(* Logix 5000 project; controller TFF vendor 1 type 14 code 107 rev 33.11; software revision 33.04; part 29 of 38 *)
(* tags used below, declared in another part *)
   Address : DINT;   // Temp Address
   BufferSteps0_Prev : STRING25;
   Config : Configuration;   // Index Array used in configuration routines
   Index : DINT;   // Index
   Index2 : DINT;   // Index
   RecipeStepLog_DateTime_Empty : STRING25;   // Empty String
   RecipeStepLog_DateTime_Log : STRING25;   // Last Date Time Received from HMI
   RecipeStepLog_DateTime_Prev : STRING25;
   RecipeStepLog_Timer : TIMER;   // RecipeStepLog WatchDog Timer
   TIME : DINT[2];
   AI01 : ALIAS FOR AnalogPoint[28];
   AI02 : ALIAS FOR AnalogPoint[29];
   AI03 : ALIAS FOR AnalogPoint[30];
   AI04 : ALIAS FOR AnalogPoint[31];
   AI104 : ALIAS FOR AnalogPoint[17];
   AI201A : ALIAS FOR AnalogPoint[10];
   AI201A_SIG : ALIAS FOR DigitalPoint[90];
   AI201B : ALIAS FOR AnalogPoint[0];
   AI202 : ALIAS FOR AnalogPoint[9];
   AI203 : ALIAS FOR AnalogPoint[11];
   AI203_SIG : ALIAS FOR DigitalPoint[91];
   AI204 : ALIAS FOR AnalogPoint[12];
   AI204_SIG : ALIAS FOR DigitalPoint[92];
   AlarmAnalog : AlarmAnalog[50];   // Analog Alarm Array
   AlarmControl : AlarmControl;   // Alarm Control
   AlarmDeviation : AlarmDeviation[20];   // Control Loop Deviation Alarm Array
   AnalogOutput : AnalogOutput[25];   // Analog Output Array
   AnalogPoint : AnalogInput[50];   // Analog Input Array
   CCPSystem : CCPSystem;   // CCP System Data
   CPU_Scanning : BOOL;   // System Scanning Flag
   DigitalOutput : BOOL[256];   // Digital Output Array these bits are sent to output cards.
   DigitalPoint : DigitalPoint[150];   // Digital Point Array
   FI101 : ALIAS FOR AnalogPoint[19];
   FI201 : ALIAS FOR AnalogPoint[2];
   FI201_SIG : ALIAS FOR DigitalPoint[93];
   FI401 : ALIAS FOR AnalogPoint[20];
   FI401_SIG : ALIAS FOR DigitalPoint[94];
   Gateway : Gateway;   // Gateway Control
   GWModbus : IO_Station;   // Status of Gateway Modbus
   HTCCollectorError : BOOL;   // Historical Data Collector Error (Set to 1 by HMI if Error)
   HTCHeartBeat : BOOL;   // Historical Data Collection heartbeat (Set to 1 by HMI Reset to 0 by PLC)
   MIX101 : ALIAS FOR AnalogPoint[14];
   Mixer : Mixer;   // Mixer config. structure
   OperatingTime : OperatingTime;
   PcToPLCHeartBeat : BOOL;   // PC to PLC communication heartbeat Set to 1 by HMI Reset to 0 by plc
   PCV101 : ALIAS FOR AnalogPoint[3];
   PCV201 : ALIAS FOR AnalogPoint[4];
   Phase0 : ALIAS FOR Phase[0];   // Phase 0
   PI001 : ALIAS FOR AnalogPoint[5];
   PI001_SIG : ALIAS FOR DigitalPoint[97];
   PI101 : ALIAS FOR AnalogPoint[6];
   PI201 : ALIAS FOR AnalogPoint[7];
   PI401 : ALIAS FOR AnalogPoint[8];
   PI601 : ALIAS FOR AnalogPoint[21];
   PI601_SIG : ALIAS FOR DigitalPoint[95];
   PLCFault : FaultRecordType;   // PLC Major Fault Record
   Rack_ACT350_WI101_200L : IO_Station;   // Status of ACT350 200L
   Rack_ACT350_WI101_500L : IO_Station;   // Status of ACT350 500L
   Rack_Murr_Node0_Smart : IO_Station;   // Status of Node 0 Smart
   Rack_Murr_Node1_TFF20 : IO_Station;   // Status of Node 1 TFF20
   Rack_Murr_Node1_TFF40 : IO_Station;   // Status of Node 1 TFF40
   Rack_Murr_Node1_TFF80 : IO_Station;   // Status of Node 1 TFF80
   RawAnalogInputArray : INT[50];   // Array of analog input raw
   RecipeStepLog_DateTime : STRING25;
   SysControl : SysControl;   // General system status and command
   Tank : TankManagement;   // Tank Management
   TCU101 : ALIAS FOR AnalogPoint[18];
   ThisSystem : SystemType;
   TI101 : ALIAS FOR AnalogPoint[13];
   TI201 : ALIAS FOR AnalogPoint[22];
   WI201 : ALIAS FOR AnalogPoint[1];
   WI201_SIG : ALIAS FOR DigitalPoint[96];
   XS011 : ALIAS FOR DigitalPoint[14];
   XS012 : ALIAS FOR DigitalPoint[15];
   YA01 : ALIAS FOR DigitalPoint[50];
   YA02 : ALIAS FOR DigitalPoint[51];
   YA03 : ALIAS FOR DigitalPoint[52];
   YA06 : ALIAS FOR DigitalPoint[55];
   YA07 : ALIAS FOR DigitalPoint[56];
   YA08 : ALIAS FOR DigitalPoint[57];
   YA09 : ALIAS FOR DigitalPoint[58];
   YA10 : ALIAS FOR DigitalPoint[59];
   YA13 : ALIAS FOR DigitalPoint[62];
   YA14 : ALIAS FOR DigitalPoint[63];
   YA15 : ALIAS FOR DigitalPoint[69];
   YA16 : ALIAS FOR DigitalPoint[70];
   YA17 : ALIAS FOR DigitalPoint[71];
   YA18 : ALIAS FOR DigitalPoint[72];
   YA41 : ALIAS FOR DigitalPoint[73];
   ZS001 : ALIAS FOR DigitalPoint[6];
   ZS002 : ALIAS FOR DigitalPoint[7];
   ZS003 : ALIAS FOR DigitalPoint[8];
   ZS004 : ALIAS FOR DigitalPoint[9];
   ZS005 : ALIAS FOR DigitalPoint[10];
   ZSDF : ALIAS FOR DigitalPoint[68];
(* Process, continued *)

ROUTINE FaultRoutine   (* ladder *)
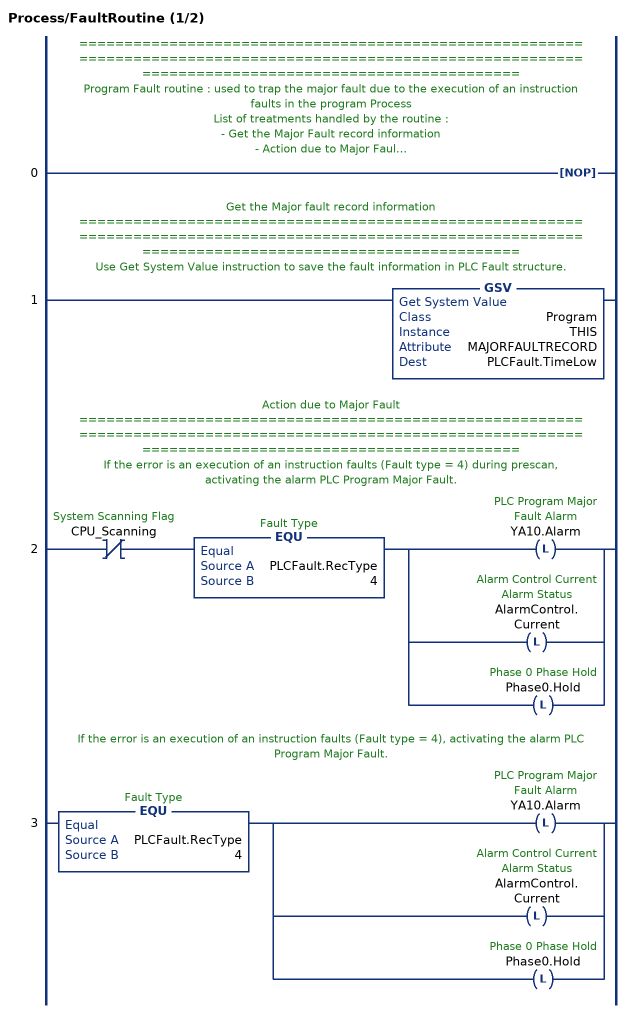
   // ==========================================================================================================================================================
   //                                                               Program Fault routine : used to trap the major fault due to the execution of an instruction faults in the program Process
   //                                                     List of treatments handled by the routine :
   //                                                          - Get the Major Fault record information
   //                                                          - Action due to Major Fault
   //                                                     -----------------------------------------------------------------------------------------------------------------------------------------------------
   //                                                     History
   // 		2019-DEC-24 - Merck - Q. Spindler - Initial version for Candidate Release 1.00.00.00.a
   // ==========================================================================================================================================================
   0: NOP();
   // Get the Major fault record information
   // ==========================================================================================================================================================
   // Use Get System Value instruction to save the fault information in PLC Fault structure.
   1: GSV(Program,THIS,MAJORFAULTRECORD,PLCFault.TimeLow);
   // Action due to Major Fault
   // ==========================================================================================================================================================
   // If the error is an execution of an instruction faults (Fault type = 4) during prescan, activating the alarm PLC Program Major Fault.
   2: XIO(CPU_Scanning)EQU(PLCFault.RecType,4)[OTL(YA10.Alarm) ,OTL(AlarmControl.Current) ,OTL(Phase0.Hold) ];
   // If the error is an execution of an instruction faults (Fault type = 4), activating the alarm PLC Program Major Fault.
   3: EQU(PLCFault.RecType,4)[OTL(YA10.Alarm) ,OTL(AlarmControl.Current) ,OTL(Phase0.Hold) ];
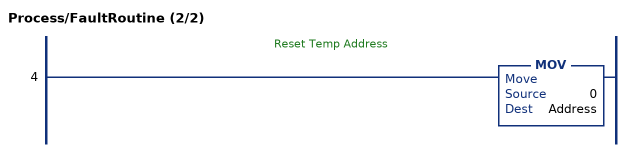
   // Reset Temp Address
   4: MOV(0,Address);
END_ROUTINE

ROUTINE Gateway   (* structured text *)
   (* ==========================================================
   	Gateway : Mapping Data to gateway communication Table
   		format of data transfered is DINT.
   		REAL type Data (Analog) must managed to convert it to DINT format with an accuracy of 3 digits (x1000 for Data sended, /1000 for Data received.
   
   	List of treatments
   		- Write to the gateway
   		- Read from the gateway
   		- Gateway wattchdog  processing
   
   -----------------------------------------------------------------------------------------------------------------------------------------------------
   	History
   		2019-DEC-24 - Merck - Q. Spindler - Initial version for Candidate Release 1.00.00.00.a
   		2020-MAR-25 - Merck - Q. Spindler - Modifications for Candidate Release 1.00.00.00.b
   					- Change Analog output indexes that caused PLC major Fault
   ============================================================*)
   
   
   
   (* Write to the gateway
   =========================================================================*)
   
   (* Send analog Point to the gateway*)
   FOR Gateway.Index := 0 TO 46 BY 1 DO
   	Gateway.Output[Gateway.Index]:= AnalogPoint[Gateway.Index].CurrentValue*1000;
   END_FOR;
   
   (* Send analog output to the gateway*)
   FOR Gateway.Index := 47 TO 58 BY 1 DO
   	Gateway.Output[Gateway.Index]:= AnalogOutput[Gateway.Index-47].ScaledValue*1000;
   END_FOR;
   
   (* Send Digital Point to the gateway*)
   FOR Gateway.Index := 0 TO 31 BY 1 DO
   	Gateway.Output[59].[Gateway.Index]:= DigitalPoint[Gateway.Index].CurrentValue;
   	Gateway.Output[60].[Gateway.Index]:= DigitalPoint[Gateway.Index+32].CurrentValue;
   	Gateway.Output[61].[Gateway.Index]:= DigitalPoint[Gateway.Index+50].SoftInput;
   	Gateway.Output[62].[Gateway.Index]:= DigitalPoint[Gateway.Index+82].SoftInput;
   END_FOR;
   
   (* Send Digital Output to the gateway *)
   FOR Gateway.Index := 0 TO 31 BY 1 DO
   	Gateway.Output[63].[Gateway.Index]:= DigitalOutput[Gateway.Index];
   	Gateway.Output[64].[Gateway.Index]:= DigitalOutput[Gateway.Index+32];
   	Gateway.Output[65].[Gateway.Index]:= DigitalOutput[Gateway.Index+64];
   END_FOR;
   
   (* Send Digital Alarm to the gateway*)
   FOR Gateway.Index := 0 TO 31 BY 1 DO
   	Gateway.Output[66].[Gateway.Index]:= DigitalPoint[Gateway.Index].Alarm;
   	Gateway.Output[67].[Gateway.Index]:= DigitalPoint[Gateway.Index+32].Alarm;
   	Gateway.Output[68].[Gateway.Index]:= DigitalPoint[Gateway.Index+64].Alarm;
   	Gateway.Output[69].[Gateway.Index]:= DigitalPoint[Gateway.Index+96].Alarm;
   END_FOR;
   
   
   (* Send Analog Alarm to the gateway*)
   FOR Gateway.Index := 70 TO 75 BY 1 DO
   	FOR Gateway.Index2 := 0 TO 31 BY 4 DO
   		Gateway.Output[Gateway.Index].[Gateway.Index2] := AlarmAnalog[(Gateway.Index2 / 4)+((Gateway.Index-70) * 8)].LOLOAlarm;
   		Gateway.Output[Gateway.Index].[Gateway.Index2 + 1] := AlarmAnalog[(Gateway.Index2 / 4)+((Gateway.Index-70) * 8)].LOAlarm;
   		Gateway.Output[Gateway.Index].[Gateway.Index2 + 2] := AlarmAnalog[(Gateway.Index2 / 4)+((Gateway.Index-70) * 8)].HIAlarm;
   		Gateway.Output[Gateway.Index].[Gateway.Index2 + 3] := AlarmAnalog[(Gateway.Index2 / 4)+((Gateway.Index-70) * 8)].HIHIAlarm;
   	END_FOR;
   END_FOR;
   
   
   (* Send Deviqtions Alarm to the gateway*)
   FOR Gateway.Index := 0 TO 15 BY 1 DO
   	Gateway.Output[76].[Gateway.Index * 2] := AlarmDeviation[Gateway.Index].HIAlarm;
   	Gateway.Output[76].[Gateway.Index * 2 + 1] := AlarmDeviation[Gateway.Index].HIHIAlarm;
   END_FOR;
   
   (* Clear unused space*)
   FOR Gateway.Index := 77 TO 81 BY 1 DO
   	Gateway.Output[Gateway.Index] := 0;
   END_FOR;
   
   
   (* Send CCP System status, system in alarm status, system in maintenance mode status to the gateway*)
   Gateway.Output[82] := CCPSystem.State;
   Gateway.Output[83].0 := AlarmControl.AlarmHigh ;
   Gateway.Output[83].1 := AlarmControl.AlarmLow ;
   Gateway.Output[83].2 := SysControl.Maintenance;
   
   (* Send Analog Action from recipe to the gateway *)
   FOR Gateway.Index := 84 TO 103 BY 1 DO
   	Gateway.Output[Gateway.Index]:= Gateway.RecipeAction_Analog[Gateway.Index-84]*1000;
   END_FOR;
   
   (* Send Digital Action from recipe to the gateway *)
   FOR Gateway.Index := 104 TO 105 BY 1 DO
   	Gateway.Output[Gateway.Index]:= Gateway.RecipeAction_Digital[Gateway.Index-104];
   END_FOR;
   
   (* Send Watchdog data to the gateway *)
   Gateway.Output[106] := Gateway.Watchdog_Out_Skid;
   Gateway.Output[107] := Gateway.Watchdog_Out_Ext;
   
   (* Data Send to the Gateway*)
   FOR Gateway.Index := 0 TO 123 BY 1 DO
   	GATEWAY:O.Data[Gateway.Index] := Gateway.Output[Gateway.Index];
   END_FOR;
   
   
   (* Read from the gateway
   =========================================================================*)
   
   (* Read from the gateway tha analog criteria for recipe *)
   FOR Gateway.Index := 0 TO 19 BY 1 DO
   		Gateway.RecipeCriteria_Analog[Gateway.Index] := Gateway.Input[Gateway.Index]/1000;
   END_FOR;
   
   (* Read from the gateway tha digital criteria for recipe *)
   FOR Gateway.Index := 20 TO 21 BY 1 DO
   		Gateway.RecipeCriteria_Digital[Gateway.Index-20] := Gateway.Input[Gateway.Index];
   END_FOR;
   
   (* Read Watchdog data from the gateway *)
   Gateway.Watchdog_In_Skid := Gateway.Input[22];
   Gateway.Watchdog_In_Ext := Gateway.Input[23];
   
   (* Data receive from the Gateway *)
   FOR Gateway.Index := 0 TO 63 BY 1 DO
   	Gateway.Input[Gateway.Index] := GATEWAY:I.Data[Gateway.Index];
   END_FOR;
   
   
   
   (* Gateway wattchdog  processing
   =========================================================================*)
   
   (* Verify if skid watchdog value receive is equal to watchdog value send previously *)
   IF Gateway.Watchdog_Out_Skid = Gateway.Watchdog_In_Skid Then
   	(* Add 1 to skid watchdog value *)
   	Gateway.Watchdog_Out_Skid := Gateway.Watchdog_Out_Skid +1;
   	(* Set to 1 YA16 soft input (alarm watchdog) *)
   	YA16.SoftInput := 1 ;
   Else
   	(* Set to 0 YA16 soft input (alarm watchdog) *)
   	YA16.SoftInput := 0 ;
   End_If;
   
   (* If skid watchdog value is greater than 9999, reset value *)
   IF Gateway.Watchdog_Out_Skid > 9999 Then
   	Gateway.Watchdog_Out_Skid := 0;
   End_IF;
   
   (* Copy external watchdog value received in the one to be sent *)
   Gateway.Watchdog_Out_Ext := Gateway.Watchdog_In_Ext;
END_ROUTINE

ROUTINE InputAnalogPoint   (* ladder *)
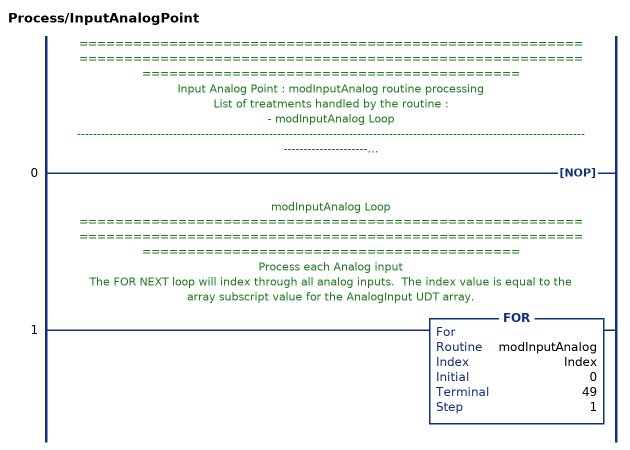
   // ==========================================================================================================================================================
   //                                                                                                             Input Analog Point : modInputAnalog routine processing
   //                                                     List of treatments handled by the routine :
   //                                                          - modInputAnalog Loop
   //                                                     -----------------------------------------------------------------------------------------------------------------------------------------------------
   //                                                     History
   // 		2019-DEC-24 - Merck - Q. Spindler - Initial version for Candidate Release 1.00.00.00.a
   // ==========================================================================================================================================================
   0: NOP();
   // modInputAnalog Loop
   // ==========================================================================================================================================================
   // Process each Analog input
   // The FOR NEXT loop will index through all analog inputs.  The index value is equal to the array subscript value for the AnalogInput UDT array.
   1: FOR(modInputAnalog,Index,0,49,1);
END_ROUTINE

ROUTINE InputAnalogRaw   (* ladder *)
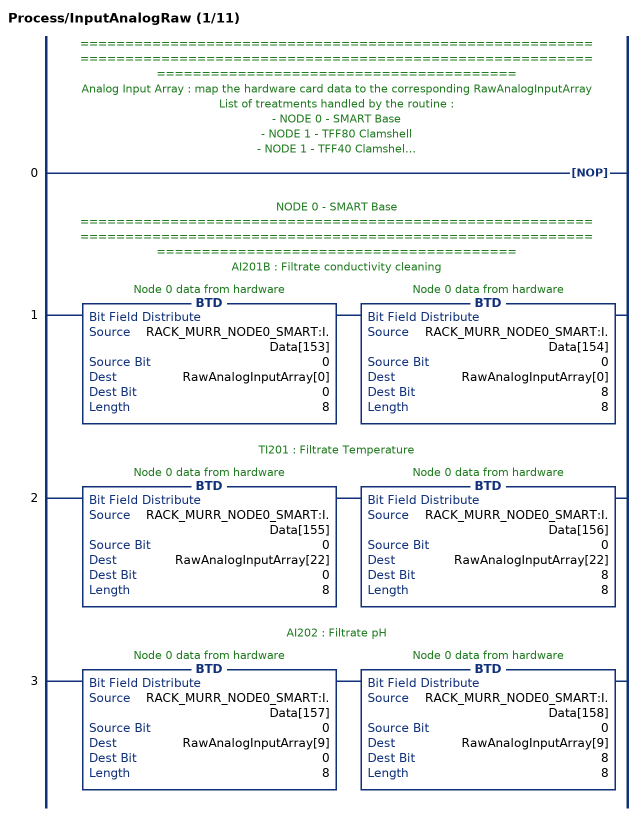
   // ==========================================================================================================================================================
   //                                                                                          Analog Input Array : map the hardware card data to the corresponding RawAnalogInputArray
   //                                                     List of treatments handled by the routine :
   //                                                    - NODE 0 - SMART Base
   //                                                         - NODE 1 - TFF80 Clamshell
   //                                                         - NODE 1 - TFF40 Clamshell
   //                                                         - NODE 1 - TFF20 Clamshell
   //                                                     -----------------------------------------------------------------------------------------------------------------------------------------------------
   //                                                     History
   // 		2019-DEC-24 - Merck - Q. Spindler - Initial version for Candidate Release 1.00.00.00.a
   //                                 2020-APR-09 - Merck - Q. Spindler - Modifications for Candidate Release 1.00.00.00.b
   //                  - Change IO address for MIX101
   //                                 2022-SEP-28 - Actemium - J. Jaekel - Modifications for Candidate Release 1.01.00.01.a
   // - Add TI201
   // ==========================================================================================================================================================
   0: NOP();
   // NODE 0 - SMART Base
   // ==========================================================================================================================================================
   // AI201B : Filtrate conductivity cleaning
   1: BTD(RACK_MURR_NODE0_SMART:I.Data[153],0,RawAnalogInputArray[0],0,8)BTD(RACK_MURR_NODE0_SMART:I.Data[154],0,RawAnalogInputArray[0],8,8);
   // TI201 : Filtrate Temperature
   2: BTD(RACK_MURR_NODE0_SMART:I.Data[155],0,RawAnalogInputArray[22],0,8)BTD(RACK_MURR_NODE0_SMART:I.Data[156],0,RawAnalogInputArray[22],8,8);
   // AI202 : Filtrate pH
   3: BTD(RACK_MURR_NODE0_SMART:I.Data[157],0,RawAnalogInputArray[9],0,8)BTD(RACK_MURR_NODE0_SMART:I.Data[158],0,RawAnalogInputArray[9],8,8);
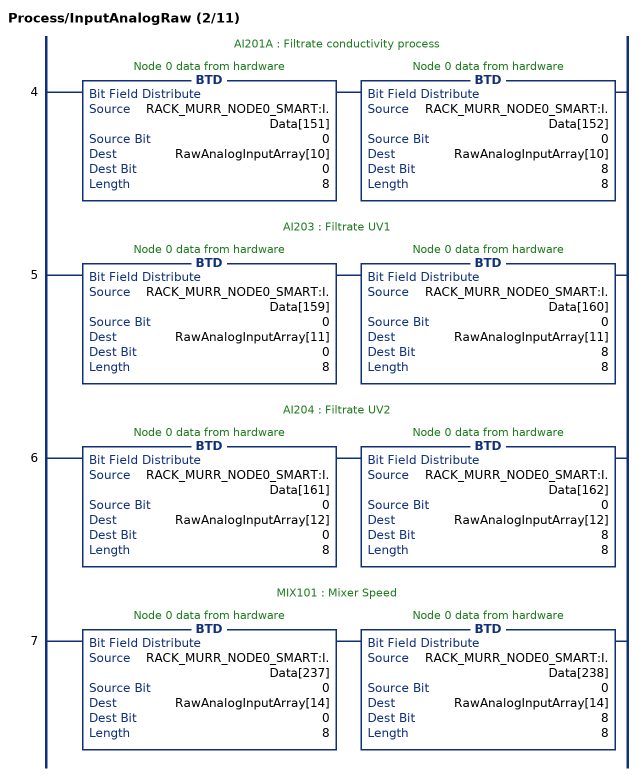
   // AI201A : Filtrate conductivity process
   4: BTD(RACK_MURR_NODE0_SMART:I.Data[151],0,RawAnalogInputArray[10],0,8)BTD(RACK_MURR_NODE0_SMART:I.Data[152],0,RawAnalogInputArray[10],8,8);
   // AI203 : Filtrate UV1
   5: BTD(RACK_MURR_NODE0_SMART:I.Data[159],0,RawAnalogInputArray[11],0,8)BTD(RACK_MURR_NODE0_SMART:I.Data[160],0,RawAnalogInputArray[11],8,8);
   // AI204 : Filtrate UV2
   6: BTD(RACK_MURR_NODE0_SMART:I.Data[161],0,RawAnalogInputArray[12],0,8)BTD(RACK_MURR_NODE0_SMART:I.Data[162],0,RawAnalogInputArray[12],8,8);
   // MIX101 : Mixer Speed
   7: BTD(RACK_MURR_NODE0_SMART:I.Data[237],0,RawAnalogInputArray[14],0,8)BTD(RACK_MURR_NODE0_SMART:I.Data[238],0,RawAnalogInputArray[14],8,8);
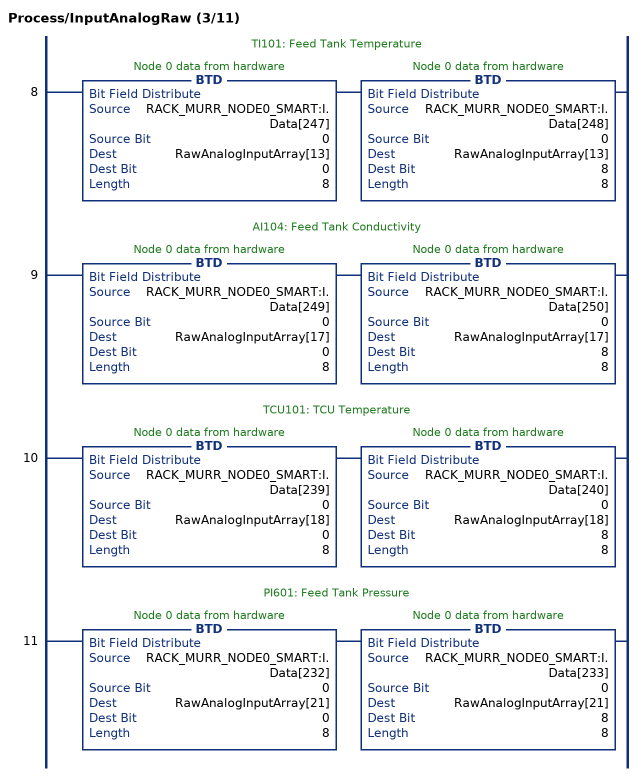
   // TI101: Feed Tank Temperature
   8: BTD(RACK_MURR_NODE0_SMART:I.Data[247],0,RawAnalogInputArray[13],0,8)BTD(RACK_MURR_NODE0_SMART:I.Data[248],0,RawAnalogInputArray[13],8,8);
   // AI104: Feed Tank Conductivity
   9: BTD(RACK_MURR_NODE0_SMART:I.Data[249],0,RawAnalogInputArray[17],0,8)BTD(RACK_MURR_NODE0_SMART:I.Data[250],0,RawAnalogInputArray[17],8,8);
   // TCU101: TCU Temperature
   10: BTD(RACK_MURR_NODE0_SMART:I.Data[239],0,RawAnalogInputArray[18],0,8)BTD(RACK_MURR_NODE0_SMART:I.Data[240],0,RawAnalogInputArray[18],8,8);
   // PI601: Feed Tank Pressure
   11: BTD(RACK_MURR_NODE0_SMART:I.Data[232],0,RawAnalogInputArray[21],0,8)BTD(RACK_MURR_NODE0_SMART:I.Data[233],0,RawAnalogInputArray[21],8,8);
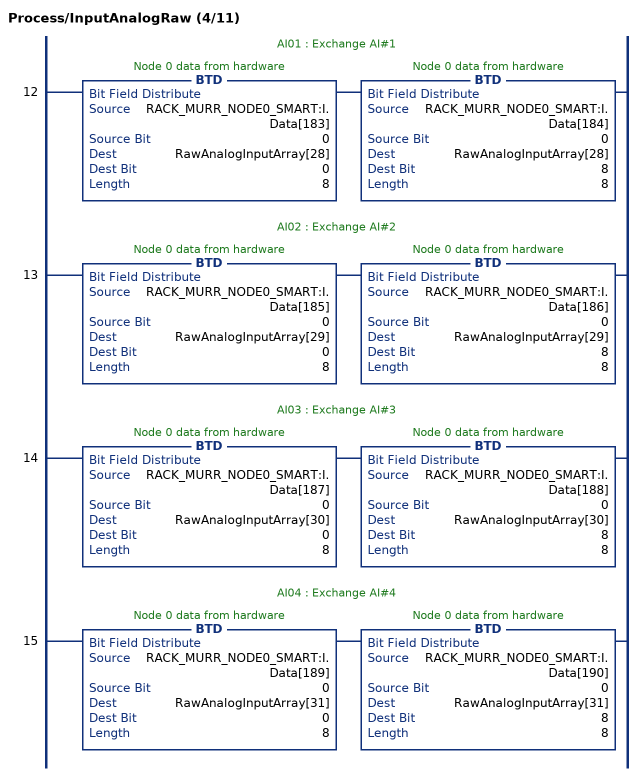
   // AI01 : Exchange AI#1
   12: BTD(RACK_MURR_NODE0_SMART:I.Data[183],0,RawAnalogInputArray[28],0,8)BTD(RACK_MURR_NODE0_SMART:I.Data[184],0,RawAnalogInputArray[28],8,8);
   // AI02 : Exchange AI#2
   13: BTD(RACK_MURR_NODE0_SMART:I.Data[185],0,RawAnalogInputArray[29],0,8)BTD(RACK_MURR_NODE0_SMART:I.Data[186],0,RawAnalogInputArray[29],8,8);
   // AI03 : Exchange AI#3
   14: BTD(RACK_MURR_NODE0_SMART:I.Data[187],0,RawAnalogInputArray[30],0,8)BTD(RACK_MURR_NODE0_SMART:I.Data[188],0,RawAnalogInputArray[30],8,8);
   // AI04 : Exchange AI#4
   15: BTD(RACK_MURR_NODE0_SMART:I.Data[189],0,RawAnalogInputArray[31],0,8)BTD(RACK_MURR_NODE0_SMART:I.Data[190],0,RawAnalogInputArray[31],8,8);
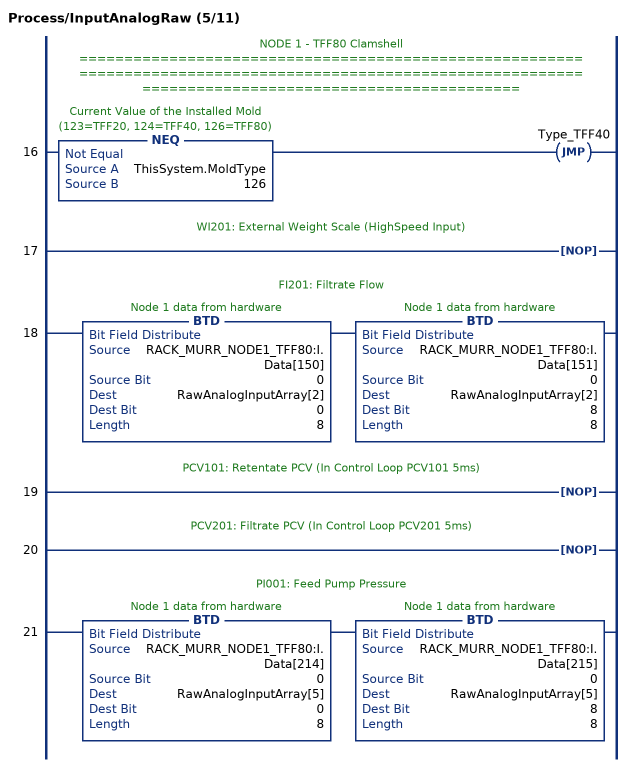
   // NODE 1 - TFF80 Clamshell
   // ==========================================================================================================================================================
   16: NEQ(ThisSystem.MoldType,126)JMP(Type_TFF40);
   // WI201: External Weight Scale (HighSpeed Input)
   17: NOP();
   // FI201: Filtrate Flow
   18: BTD(RACK_MURR_NODE1_TFF80:I.Data[150],0,RawAnalogInputArray[2],0,8)BTD(RACK_MURR_NODE1_TFF80:I.Data[151],0,RawAnalogInputArray[2],8,8);
   // PCV101: Retentate PCV (In Control Loop PCV101 5ms)
   19: NOP();
   // PCV201: Filtrate PCV (In Control Loop PCV201 5ms)
   20: NOP();
   // PI001: Feed Pump Pressure
   21: BTD(RACK_MURR_NODE1_TFF80:I.Data[214],0,RawAnalogInputArray[5],0,8)BTD(RACK_MURR_NODE1_TFF80:I.Data[215],0,RawAnalogInputArray[5],8,8);
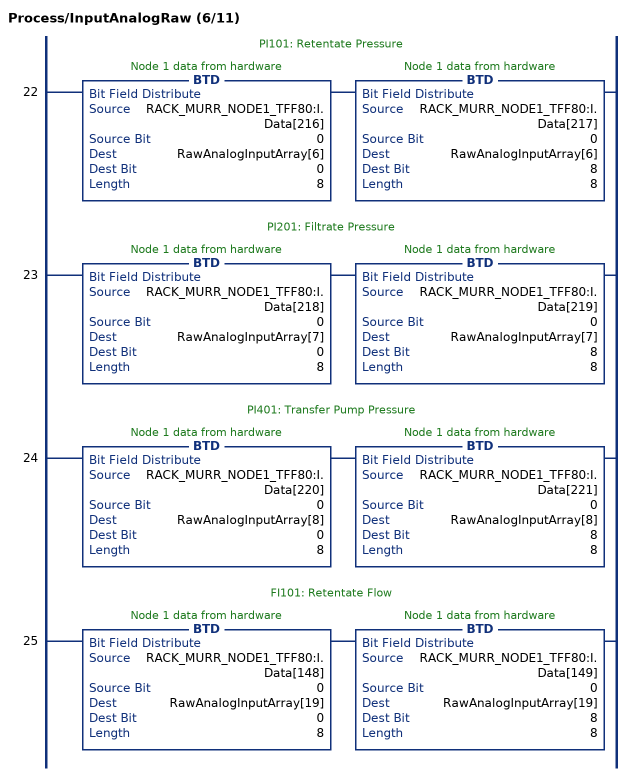
   // PI101: Retentate Pressure
   22: BTD(RACK_MURR_NODE1_TFF80:I.Data[216],0,RawAnalogInputArray[6],0,8)BTD(RACK_MURR_NODE1_TFF80:I.Data[217],0,RawAnalogInputArray[6],8,8);
   // PI201: Filtrate Pressure
   23: BTD(RACK_MURR_NODE1_TFF80:I.Data[218],0,RawAnalogInputArray[7],0,8)BTD(RACK_MURR_NODE1_TFF80:I.Data[219],0,RawAnalogInputArray[7],8,8);
   // PI401: Transfer Pump Pressure
   24: BTD(RACK_MURR_NODE1_TFF80:I.Data[220],0,RawAnalogInputArray[8],0,8)BTD(RACK_MURR_NODE1_TFF80:I.Data[221],0,RawAnalogInputArray[8],8,8);
   // FI101: Retentate Flow
   25: BTD(RACK_MURR_NODE1_TFF80:I.Data[148],0,RawAnalogInputArray[19],0,8)BTD(RACK_MURR_NODE1_TFF80:I.Data[149],0,RawAnalogInputArray[19],8,8);
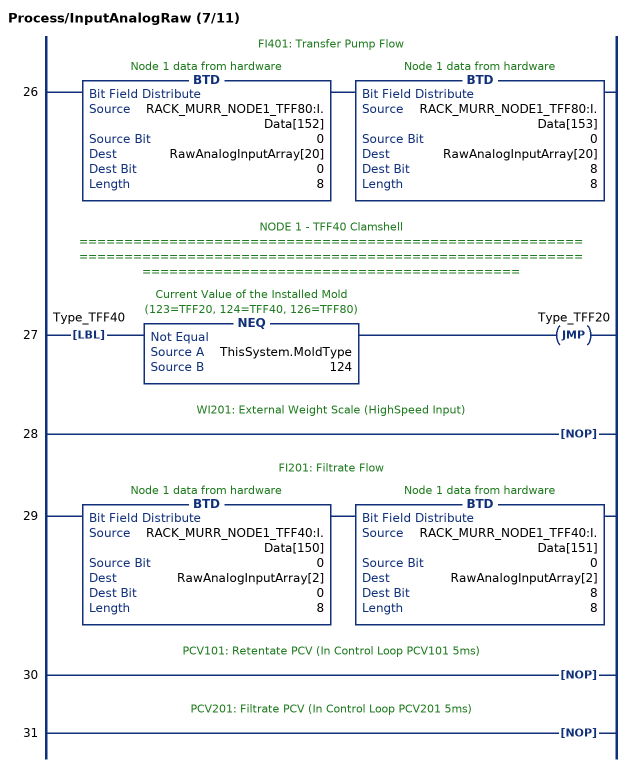
   // FI401: Transfer Pump Flow
   26: BTD(RACK_MURR_NODE1_TFF80:I.Data[152],0,RawAnalogInputArray[20],0,8)BTD(RACK_MURR_NODE1_TFF80:I.Data[153],0,RawAnalogInputArray[20],8,8);
   // NODE 1 - TFF40 Clamshell
   // ==========================================================================================================================================================
   27: LBL(Type_TFF40)NEQ(ThisSystem.MoldType,124)JMP(Type_TFF20);
   // WI201: External Weight Scale (HighSpeed Input)
   28: NOP();
   // FI201: Filtrate Flow
   29: BTD(RACK_MURR_NODE1_TFF40:I.Data[150],0,RawAnalogInputArray[2],0,8)BTD(RACK_MURR_NODE1_TFF40:I.Data[151],0,RawAnalogInputArray[2],8,8);
   // PCV101: Retentate PCV (In Control Loop PCV101 5ms)
   30: NOP();
   // PCV201: Filtrate PCV (In Control Loop PCV201 5ms)
   31: NOP();
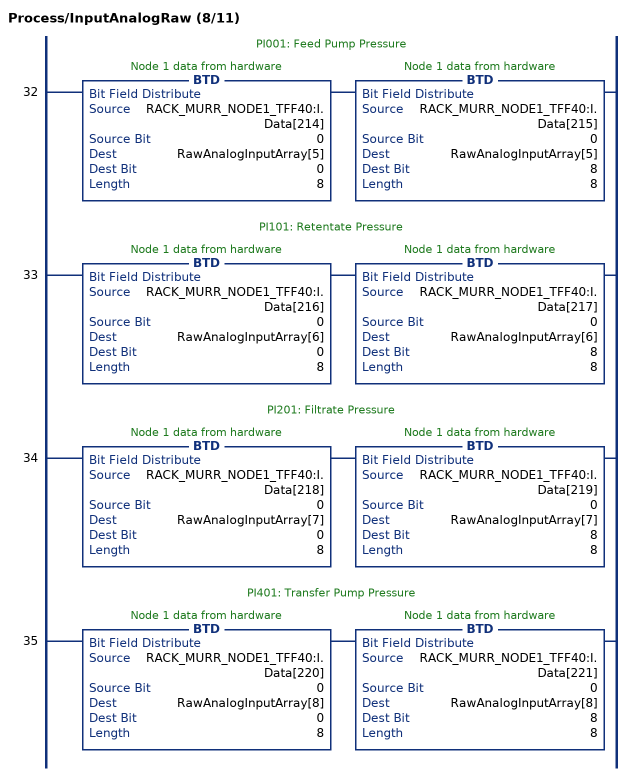
   // PI001: Feed Pump Pressure
   32: BTD(RACK_MURR_NODE1_TFF40:I.Data[214],0,RawAnalogInputArray[5],0,8)BTD(RACK_MURR_NODE1_TFF40:I.Data[215],0,RawAnalogInputArray[5],8,8);
   // PI101: Retentate Pressure
   33: BTD(RACK_MURR_NODE1_TFF40:I.Data[216],0,RawAnalogInputArray[6],0,8)BTD(RACK_MURR_NODE1_TFF40:I.Data[217],0,RawAnalogInputArray[6],8,8);
   // PI201: Filtrate Pressure
   34: BTD(RACK_MURR_NODE1_TFF40:I.Data[218],0,RawAnalogInputArray[7],0,8)BTD(RACK_MURR_NODE1_TFF40:I.Data[219],0,RawAnalogInputArray[7],8,8);
   // PI401: Transfer Pump Pressure
   35: BTD(RACK_MURR_NODE1_TFF40:I.Data[220],0,RawAnalogInputArray[8],0,8)BTD(RACK_MURR_NODE1_TFF40:I.Data[221],0,RawAnalogInputArray[8],8,8);
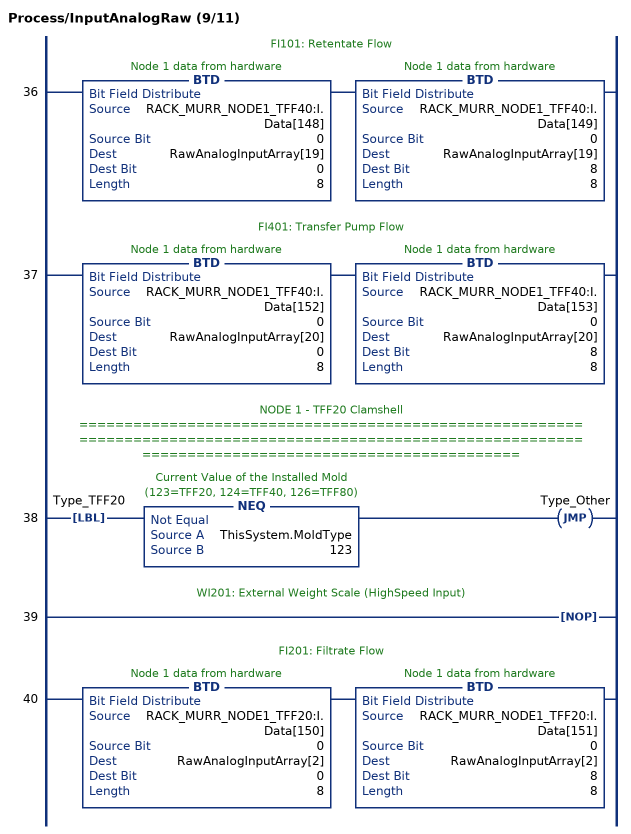
   // FI101: Retentate Flow
   36: BTD(RACK_MURR_NODE1_TFF40:I.Data[148],0,RawAnalogInputArray[19],0,8)BTD(RACK_MURR_NODE1_TFF40:I.Data[149],0,RawAnalogInputArray[19],8,8);
   // FI401: Transfer Pump Flow
   37: BTD(RACK_MURR_NODE1_TFF40:I.Data[152],0,RawAnalogInputArray[20],0,8)BTD(RACK_MURR_NODE1_TFF40:I.Data[153],0,RawAnalogInputArray[20],8,8);
   // NODE 1 - TFF20 Clamshell
   // ==========================================================================================================================================================
   38: LBL(Type_TFF20)NEQ(ThisSystem.MoldType,123)JMP(Type_Other);
   // WI201: External Weight Scale (HighSpeed Input)
   39: NOP();
   // FI201: Filtrate Flow
   40: BTD(RACK_MURR_NODE1_TFF20:I.Data[150],0,RawAnalogInputArray[2],0,8)BTD(RACK_MURR_NODE1_TFF20:I.Data[151],0,RawAnalogInputArray[2],8,8);
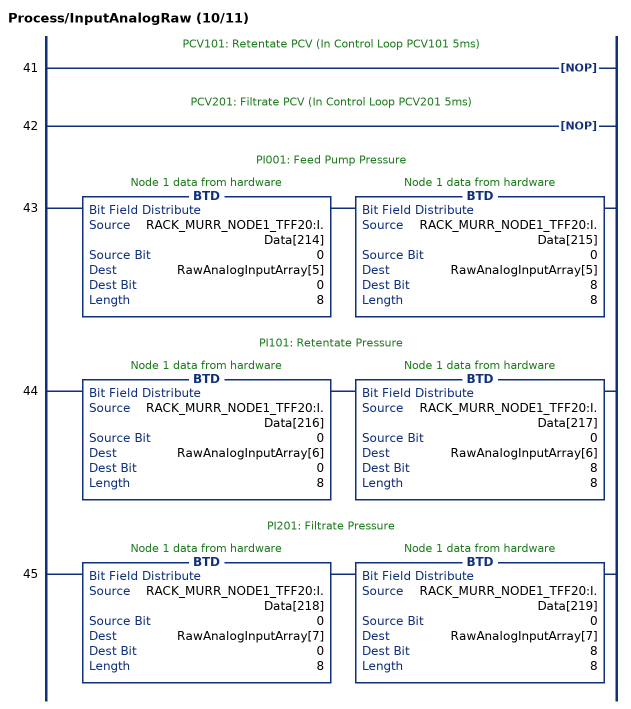
   // PCV101: Retentate PCV (In Control Loop PCV101 5ms)
   41: NOP();
   // PCV201: Filtrate PCV (In Control Loop PCV201 5ms)
   42: NOP();
   // PI001: Feed Pump Pressure
   43: BTD(RACK_MURR_NODE1_TFF20:I.Data[214],0,RawAnalogInputArray[5],0,8)BTD(RACK_MURR_NODE1_TFF20:I.Data[215],0,RawAnalogInputArray[5],8,8);
   // PI101: Retentate Pressure
   44: BTD(RACK_MURR_NODE1_TFF20:I.Data[216],0,RawAnalogInputArray[6],0,8)BTD(RACK_MURR_NODE1_TFF20:I.Data[217],0,RawAnalogInputArray[6],8,8);
   // PI201: Filtrate Pressure
   45: BTD(RACK_MURR_NODE1_TFF20:I.Data[218],0,RawAnalogInputArray[7],0,8)BTD(RACK_MURR_NODE1_TFF20:I.Data[219],0,RawAnalogInputArray[7],8,8);
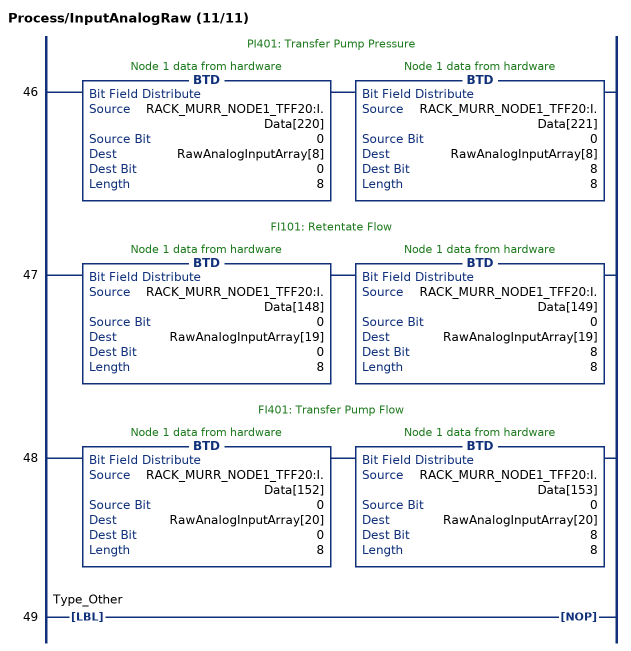
   // PI401: Transfer Pump Pressure
   46: BTD(RACK_MURR_NODE1_TFF20:I.Data[220],0,RawAnalogInputArray[8],0,8)BTD(RACK_MURR_NODE1_TFF20:I.Data[221],0,RawAnalogInputArray[8],8,8);
   // FI101: Retentate Flow
   47: BTD(RACK_MURR_NODE1_TFF20:I.Data[148],0,RawAnalogInputArray[19],0,8)BTD(RACK_MURR_NODE1_TFF20:I.Data[149],0,RawAnalogInputArray[19],8,8);
   // FI401: Transfer Pump Flow
   48: BTD(RACK_MURR_NODE1_TFF20:I.Data[152],0,RawAnalogInputArray[20],0,8)BTD(RACK_MURR_NODE1_TFF20:I.Data[153],0,RawAnalogInputArray[20],8,8);
   49: LBL(Type_Other)NOP();
END_ROUTINE

ROUTINE InputDigitalPoint   (* ladder *)
// Digital Point Routine
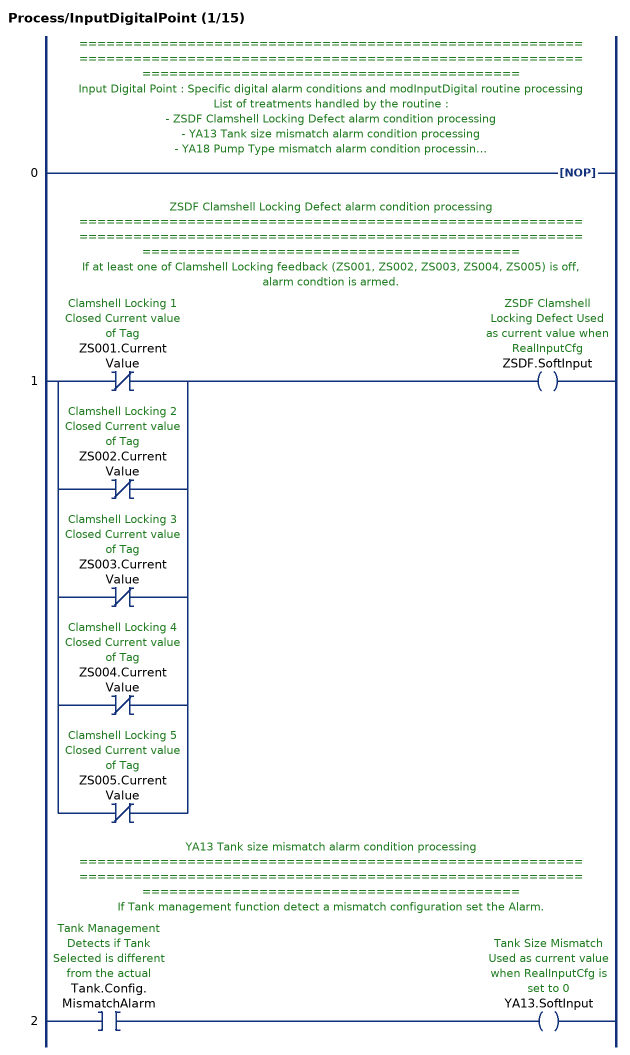
   // ==========================================================================================================================================================
   //                                                                                   Input Digital Point : Specific digital alarm conditions and modInputDigital routine processing
   //                                                     List of treatments handled by the routine :
   //                                                          - ZSDF Clamshell Locking Defect alarm condition processing
   //                                                          - YA13 Tank size mismatch alarm condition processing
   //                                                          - YA18 Pump Type mismatch alarm condition processing
   //                                                          - YA03 Historical data collection failure alarm condition processing
   //                                                          - YA01 PC to PLC com. failure alarm condition processing
   //                                                          - YA02 CCP Runtime com. failure alarm condition processing
   //                                                          - YA14 SQL Write failure alarm condition processing
   //                                                          - Node 0 communication failure and internal defect (YA06 and YA07)
   //                                                          - Node 1 communication failure and internal defect (YA08 and YA09)
   //                                                          - ACT350 communication failure (YA15)
   //                                                          - Operating Time Exceeded (YA41)
   //                                                          - Analog Signal Failure
   //                                                          - modInputDigital Loop
   //                                                     -----------------------------------------------------------------------------------------------------------------------------------------------------
   //                                                     History
   // 		2019-DEC-24 - Merck - Q. Spindler - Initial version for Candidate Release 1.00.00.00.a
   // 		2020-APR-06 - Merck - Q. Spindler - Modifications for Candidate Release 1.00.00.00.b
   //                                                             - Trigger pressure signal failure when the raw value equal to the RawMax
   // 		2020-JUN-09 - Merck - Q. Spindler - Modifications for Candidate Release 1.00.00.00.c
   //                                                             - Change Alarm condition for YA07 and YA09, internal defect dont trigger if the Node is not connected
   // - Change YA14 Alarm condition processing to add HMI Watchdog
   // 		2021-OCT-26 - Merck - Q. Spindler - Modifications for Candidate Release 1.01.00.00.a
   // - Add HTC Collector Error in the YA03 alarm conditions
   //   - Add Operating Time Exceeded (YA41)
   // 		2022-SEP-26 - Actemium - J. Jaekel - Modifications for Candidate Release 1.01.00.01.a
   // - Add TI201 signal failure
   // ==========================================================================================================================================================
   0: NOP();
   // ZSDF Clamshell Locking Defect alarm condition processing
   // ==========================================================================================================================================================
   // If at least one of Clamshell Locking feedback (ZS001, ZS002, ZS003, ZS004, ZS005) is off, alarm condtion is armed.
   1: [XIO(ZS001.CurrentValue) ,XIO(ZS002.CurrentValue) ,XIO(ZS003.CurrentValue) ,XIO(ZS004.CurrentValue) ,XIO(ZS005.CurrentValue) ]OTE(ZSDF.SoftInput);
   // YA13 Tank size mismatch alarm condition processing
   // ==========================================================================================================================================================
   // If Tank management function detect a mismatch configuration set the Alarm.
   2: XIC(Tank.Config.MismatchAlarm)OTE(YA13.SoftInput);
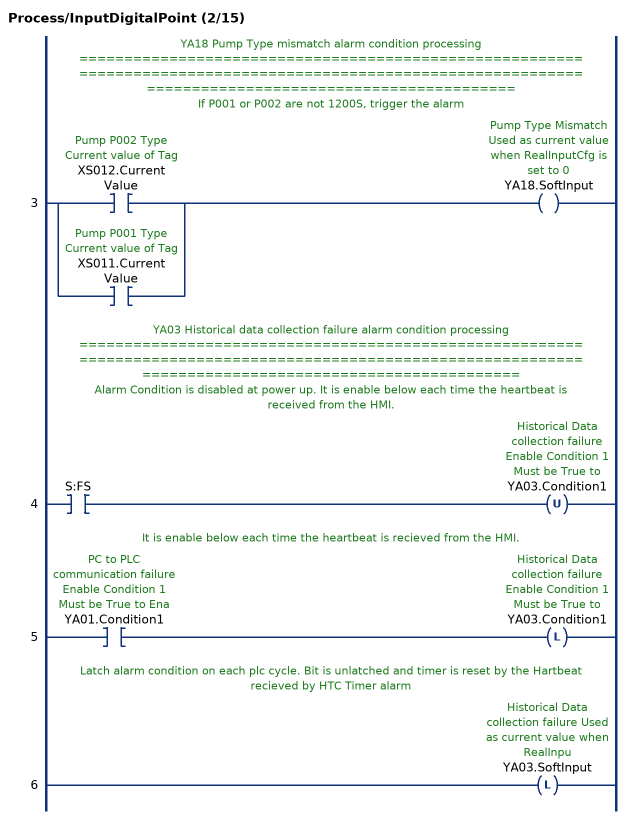
   // YA18 Pump Type mismatch alarm condition processing
   // =========================================================================================================================================================
   // If P001 or P002 are not 1200S, trigger the alarm
   3: [XIC(XS012.CurrentValue) ,XIC(XS011.CurrentValue) ]OTE(YA18.SoftInput);
   // YA03 Historical data collection failure alarm condition processing
   // ==========================================================================================================================================================
   // Alarm Condition is disabled at power up. It is enable below each time the heartbeat is received from the HMI.
   4: XIC(S:FS)OTU(YA03.Condition1);
   // It is enable below each time the heartbeat is recieved from the HMI.
   5: XIC(YA01.Condition1)OTL(YA03.Condition1);
   // Latch alarm condition on each plc cycle. Bit is unlatched and timer is reset by the Hartbeat recieved by HTC Timer alarm
   6: OTL(YA03.SoftInput);
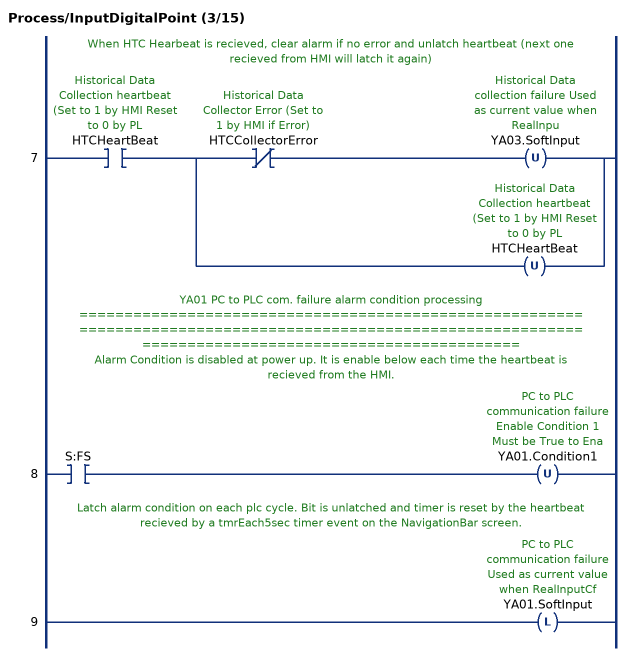
   // When HTC Hearbeat is recieved, clear alarm if no error and unlatch heartbeat (next one recieved from HMI will latch it again)
   7: XIC(HTCHeartBeat)[XIO(HTCCollectorError) OTU(YA03.SoftInput) ,OTU(HTCHeartBeat) ];
   // YA01 PC to PLC com. failure alarm condition processing
   // ==========================================================================================================================================================
   // Alarm Condition is disabled at power up. It is enable below each time the heartbeat is recieved from the HMI.
   8: XIC(S:FS)OTU(YA01.Condition1);
   // Latch alarm condition on each plc cycle. Bit is unlatched and timer is reset by the heartbeat recieved by a tmrEach5sec timer event on the NavigationBar screen.
   9: OTL(YA01.SoftInput);
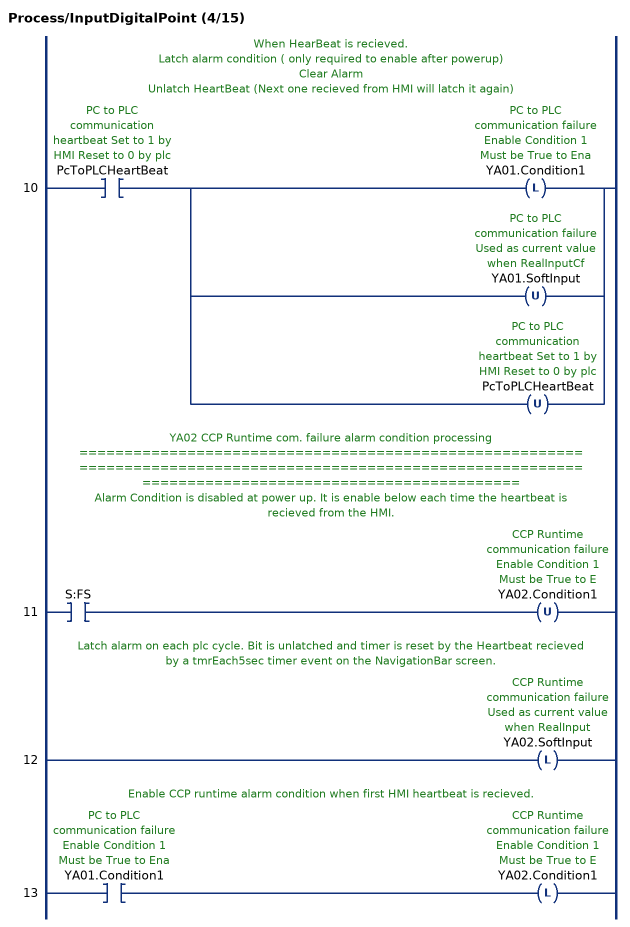
   // When HearBeat is recieved.
   //         Latch alarm condition ( only required to enable after powerup)
   //         Clear Alarm
   //        Unlatch HeartBeat (Next one recieved from HMI will latch it again)
   10: XIC(PcToPLCHeartBeat)[OTL(YA01.Condition1) ,OTU(YA01.SoftInput) ,OTU(PcToPLCHeartBeat) ];
   // YA02 CCP Runtime com. failure alarm condition processing
   // ==========================================================================================================================================================
   // Alarm Condition is disabled at power up. It is enable below each time the heartbeat is recieved from the HMI.
   11: XIC(S:FS)OTU(YA02.Condition1);
   // Latch alarm on each plc cycle. Bit is unlatched and timer is reset by the Heartbeat recieved by a tmrEach5sec timer event on the NavigationBar screen.
   12: OTL(YA02.SoftInput);
   // Enable CCP runtime alarm condition when first HMI heartbeat is recieved.
   13: XIC(YA01.Condition1)OTL(YA02.Condition1);
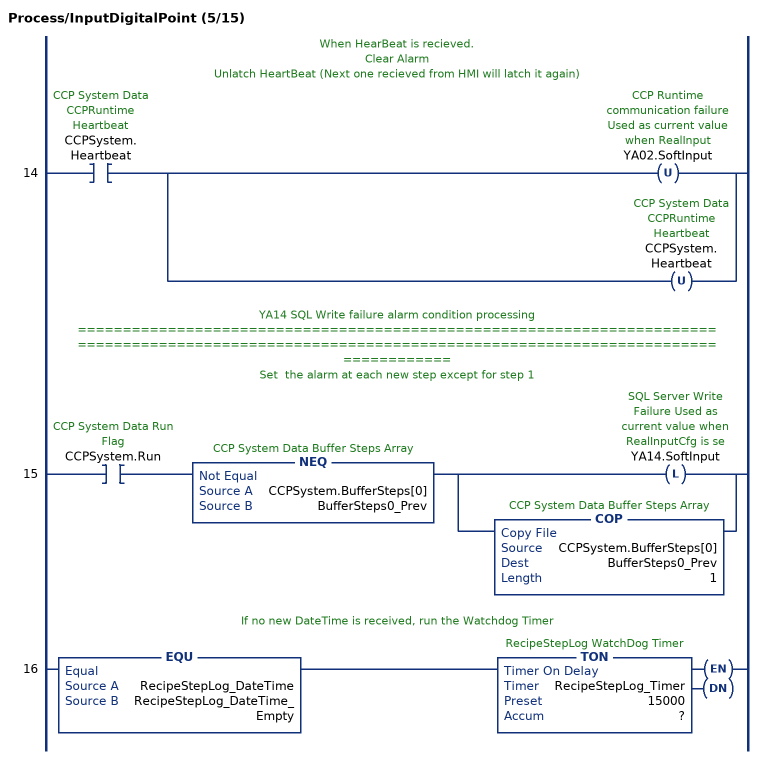
   // When HearBeat is recieved.
   //         Clear Alarm
   //        Unlatch HeartBeat (Next one recieved from HMI will latch it again)
   14: XIC(CCPSystem.Heartbeat)[OTU(YA02.SoftInput) ,OTU(CCPSystem.Heartbeat) ];
   // YA14 SQL Write failure alarm condition processing
   // ==========================================================================================================================================================
   // Set  the alarm at each new step except for step 1
   15: XIC(CCPSystem.Run)NEQ(CCPSystem.BufferSteps[0],BufferSteps0_Prev)[OTL(YA14.SoftInput) ,COP(CCPSystem.BufferSteps[0],BufferSteps0_Prev,1) ];
   // If no new DateTime is received, run the Watchdog Timer
   16: EQU(RecipeStepLog_DateTime,RecipeStepLog_DateTime_Empty)TON(RecipeStepLog_Timer,?,?);
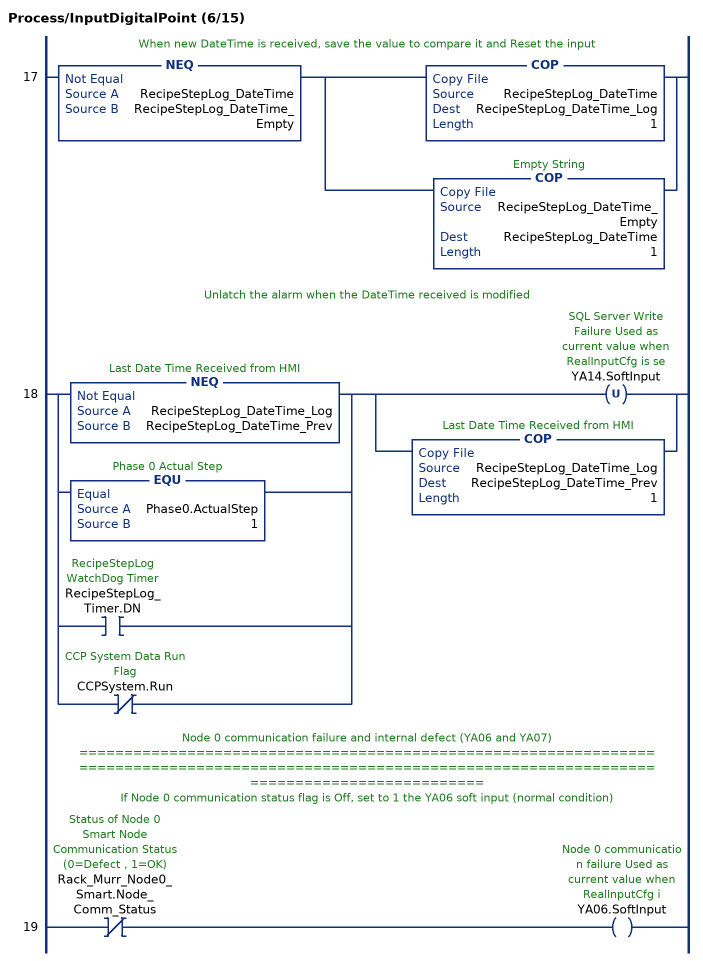
   // When new DateTime is received, save the value to compare it and Reset the input
   17: NEQ(RecipeStepLog_DateTime,RecipeStepLog_DateTime_Empty)[COP(RecipeStepLog_DateTime,RecipeStepLog_DateTime_Log,1) ,COP(RecipeStepLog_DateTime_Empty,RecipeStepLog_DateTime,1) ];
   // Unlatch the alarm when the DateTime received is modified
   18: [NEQ(RecipeStepLog_DateTime_Log,RecipeStepLog_DateTime_Prev) ,EQU(Phase0.ActualStep,1) ,XIC(RecipeStepLog_Timer.DN) ,XIO(CCPSystem.Run) ][OTU(YA14.SoftInput) ,COP(RecipeStepLog_DateTime_Log,RecipeStepLog_DateTime_Prev,1) ];
   // Node 0 communication failure and internal defect (YA06 and YA07)
   // ==========================================================================================================================================================
   // If Node 0 communication status flag is Off, set to 1 the YA06 soft input (normal condition)
   19: XIO(Rack_Murr_Node0_Smart.Node_Comm_Status)OTE(YA06.SoftInput);
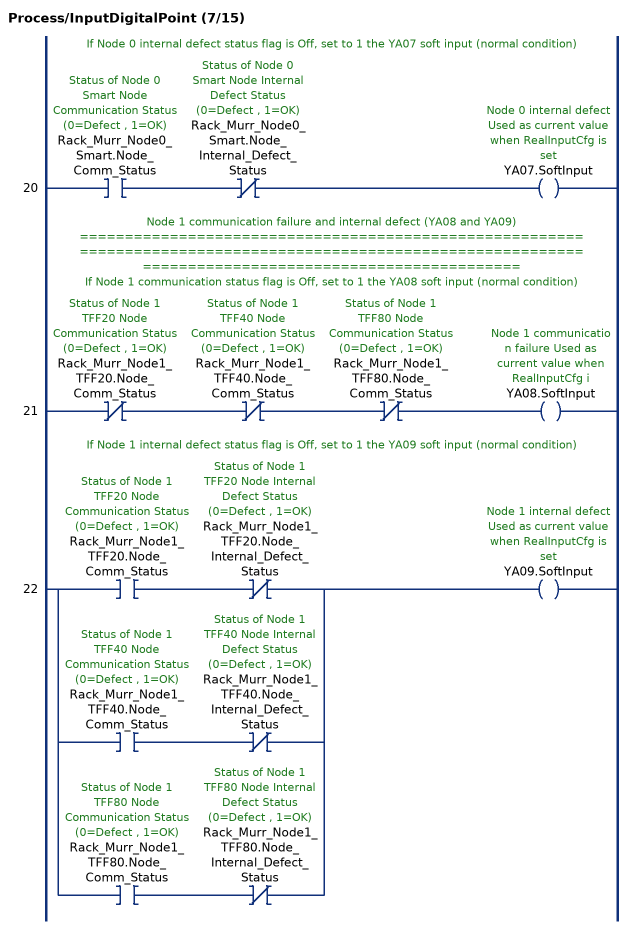
   // If Node 0 internal defect status flag is Off, set to 1 the YA07 soft input (normal condition)
   20: XIC(Rack_Murr_Node0_Smart.Node_Comm_Status)XIO(Rack_Murr_Node0_Smart.Node_Internal_Defect_Status)OTE(YA07.SoftInput);
   // Node 1 communication failure and internal defect (YA08 and YA09)
   // ==========================================================================================================================================================
   // If Node 1 communication status flag is Off, set to 1 the YA08 soft input (normal condition)
   21: XIO(Rack_Murr_Node1_TFF20.Node_Comm_Status)XIO(Rack_Murr_Node1_TFF40.Node_Comm_Status)XIO(Rack_Murr_Node1_TFF80.Node_Comm_Status)OTE(YA08.SoftInput);
   // If Node 1 internal defect status flag is Off, set to 1 the YA09 soft input (normal condition)
   22: [XIC(Rack_Murr_Node1_TFF20.Node_Comm_Status) XIO(Rack_Murr_Node1_TFF20.Node_Internal_Defect_Status) ,XIC(Rack_Murr_Node1_TFF40.Node_Comm_Status) XIO(Rack_Murr_Node1_TFF40.Node_Internal_Defect_Status) ,XIC(Rack_Murr_Node1_TFF80.Node_Comm_Status) XIO(Rack_Murr_Node1_TFF80.Node_Internal_Defect_Status) ]OTE(YA09.SoftInput);
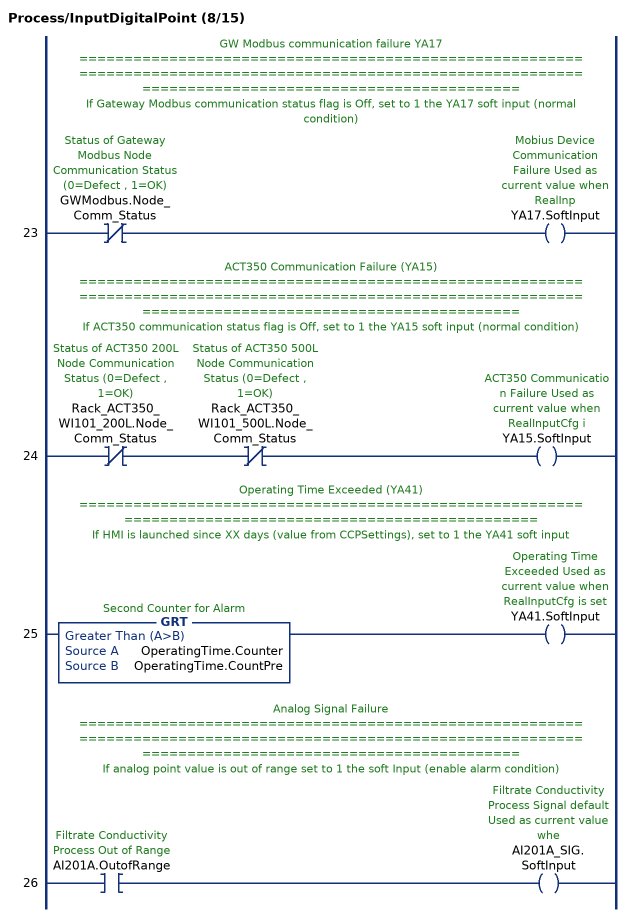
   // GW Modbus communication failure YA17
   // ==========================================================================================================================================================
   // If Gateway Modbus communication status flag is Off, set to 1 the YA17 soft input (normal condition)
   23: XIO(GWModbus.Node_Comm_Status)OTE(YA17.SoftInput);
   // ACT350 Communication Failure (YA15)
   // ==========================================================================================================================================================
   // If ACT350 communication status flag is Off, set to 1 the YA15 soft input (normal condition)
   24: XIO(Rack_ACT350_WI101_200L.Node_Comm_Status)XIO(Rack_ACT350_WI101_500L.Node_Comm_Status)OTE(YA15.SoftInput);
   // Operating Time Exceeded (YA41)
   // ======================================================================================================
   // If HMI is launched since XX days (value from CCPSettings), set to 1 the YA41 soft input
   25: GRT(OperatingTime.Counter,OperatingTime.CountPre)OTE(YA41.SoftInput);
   // Analog Signal Failure
   // ==========================================================================================================================================================
   // If analog point value is out of range set to 1 the soft Input (enable alarm condition)
   26: XIC(AI201A.OutofRange)OTE(AI201A_SIG.SoftInput);
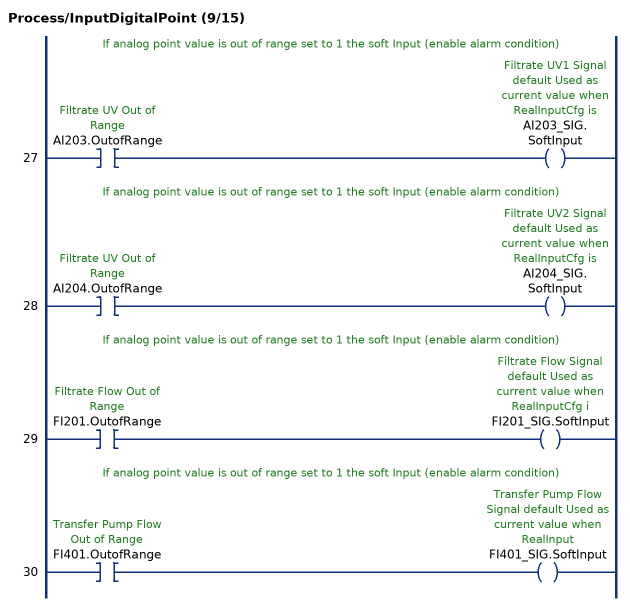
   // If analog point value is out of range set to 1 the soft Input (enable alarm condition)
   27: XIC(AI203.OutofRange)OTE(AI203_SIG.SoftInput);
   // If analog point value is out of range set to 1 the soft Input (enable alarm condition)
   28: XIC(AI204.OutofRange)OTE(AI204_SIG.SoftInput);
   // If analog point value is out of range set to 1 the soft Input (enable alarm condition)
   29: XIC(FI201.OutofRange)OTE(FI201_SIG.SoftInput);
   // If analog point value is out of range set to 1 the soft Input (enable alarm condition)
   30: XIC(FI401.OutofRange)OTE(FI401_SIG.SoftInput);
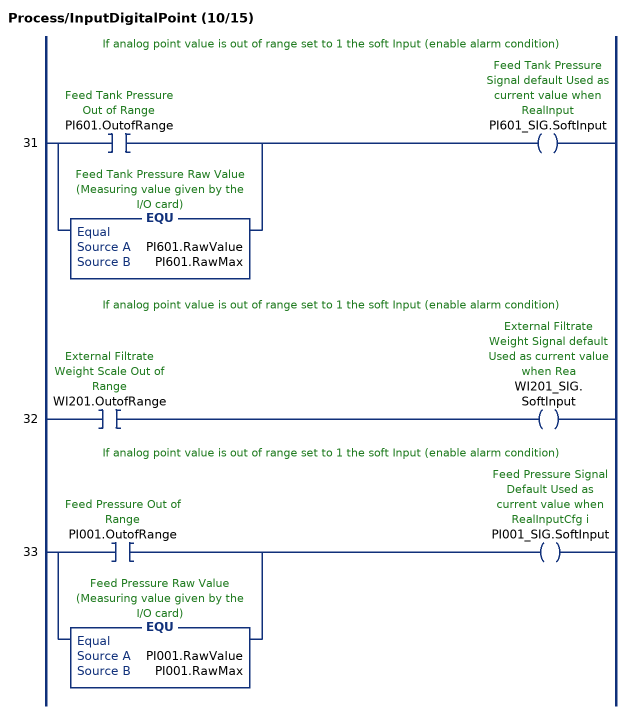
   // If analog point value is out of range set to 1 the soft Input (enable alarm condition)
   31: [XIC(PI601.OutofRange) ,EQU(PI601.RawValue,PI601.RawMax) ]OTE(PI601_SIG.SoftInput);
   // If analog point value is out of range set to 1 the soft Input (enable alarm condition)
   32: XIC(WI201.OutofRange)OTE(WI201_SIG.SoftInput);
   // If analog point value is out of range set to 1 the soft Input (enable alarm condition)
   33: [XIC(PI001.OutofRange) ,EQU(PI001.RawValue,PI001.RawMax) ]OTE(PI001_SIG.SoftInput);
